TYPE ST_IsoMon_HMI_Interface :
STRUCT
	HMIbaseDevice		: ST_Device_HMI_Interface; 
	ocmdTripReset		: BOOL;
	ocmdTest			: BOOL;
	stsDeviceAlarm		: BOOL;
	stsDeviceWarning	: BOOL;
END_STRUCT
END_TYPE

(* stored: Version 1.1.0.1
   DUT ST_IsoMon_HMI_Interface: Id {24cf9de1-fd06-492a-99f2-130270290411} *)
